Fanuc KAREL source: KO00050.KL

PROGRAM KO00050
%NOLOCKGROUP
%ENVIRONMENT MIR
VAR
  P1: XYZWPR
  P2: POSITION
  F: BOOLEAN
  OUT: XYZWPR
BEGIN
  F = TRUE
  OUT = MIRROR(P1, P2, F)
END KO00050
